(*
SPDX-FileCopyrightText: © 2026 Oleksandr Tiutyk <trofimich@gmail.com>
SPDX-License-Identifier: MIT
License: https://opensource.org/license/mit
*)

(*!
<summary>Beckhoff EL5152 32-bit incremental encoder channel without a latch.</summary>
<description>
Combines a latch-free 32-bit counter input with the 16-bit control word and 32-bit counter preset.
Select the 32-bit main PDOs for the corresponding EL5152 channel; optional period/frequency PDOs are separate.
Link input and output fields individually; the aggregate is not a packed EtherCAT packet.
Use one owner task; externally synchronize other access. Copies store data without creating hardware links.
When used for I/O, link located fields or their containing buffers to the matching selected PDOs.
The record is not a packed wire buffer; compiler padding is not part of the device specification.
Unlinked/default values do not prove valid I/O. The caller evaluates bus/channel validity before use.
Use one owner task per instance and externally synchronize other access; multi-field snapshots are not atomic.
Copies store data without creating hardware links. Keep borrowed field references valid while consumers are bound.
This passive record performs no validation, synchronization, configuration or protocol advancement.
</description>
*)
TYPE INCREMENTAL_ENCODER_COUNTER_CHANNEL :
STRUCT
	In : INCREMENTAL_ENCODER_COUNTER_INPUT_CHANNEL;
	Out : INCREMENTAL_ENCODER_OUTPUT_CHANNEL;
END_STRUCT
END_TYPE

(* stored: Version 1.1.0.1
   DUT INCREMENTAL_ENCODER_COUNTER_CHANNEL: Id {d7112403-e8dc-4964-a81d-53b6ece24076} *)
